(* IEC 61131-3 sources: PLC_I/plc/tests, 6 files *)

(* ---- 程序_气缸自测.st ---- *)
(* 离线IEC扫描自测：放入周期任务，等待b完成，w失败=0才通过。
   不连接物理输出。TON时间证据要求在目标PLC/官方模拟运行，源码测试不能替代。 *)
PROGRAM 程序_气缸自测
VAR
    fb : 功能块_气缸;
    fb原点 : 功能块_气缸;
    ui阶段 : UINT;
    w失败 : WORD;
    b完成 : BOOL;
    t等待 : TON;
    st配置 : 结构体_配置;
    fb调度 : 功能块_气缸调度;
    st运行时 : 结构体_运行时;
    lw原绑定 : LWORD;
    i : UINT;
    udi夹紧请求号 : UDINT; (* 业务示例：保存 Cy动点(Cy夹紧) 返回值 *)
END_VAR
CASE ui阶段 OF
0:
    fb(Execute := FALSE, Token := 0, Code := 0, HasWorkSensor := FALSE, HasOriginSensor := FALSE,
        DelayMs := 20, HomeDelayMs := 30, TimeoutMs := 500, ValveType := 3, HardEstop := FALSE, CancelMode := 0);
    IF fb.AtWork OR fb.AtOrigin OR (fb.DoneToken <> 0) THEN w失败 := 1; END_IF;
    ui阶段 := 1;
1:
    fb(Execute := TRUE, Token := 1, Code := 40);
    IF NOT fb.WorkOutput OR fb.OriginOutput THEN w失败 := 2; END_IF;
    IF fb.DoneToken = 1 THEN ui阶段 := 2; END_IF;
2:
    (* Execute连续TRUE，下一扫描新token仍触发反向请求。 *)
    fb(Execute := TRUE, Token := 2, Code := 41);
    IF fb.WorkOutput OR NOT fb.OriginOutput OR fb.AtWork OR (fb.DoneToken <> 0) THEN w失败 := 3; END_IF;
    ui阶段 := 3;
3:
    fb(Execute := FALSE);
    IF fb.DoneToken = 2 THEN
        IF fb.OriginOutput OR NOT fb.AtOrigin THEN w失败 := 4; END_IF;
        ui阶段 := 4;
    END_IF;
4:
    fb(Execute := TRUE, Token := 3, Code := 40);
    ui阶段 := 5;
5:
    fb(Execute := FALSE, CancelMode := 1);
    IF NOT fb.WorkOutput OR fb.Moving OR fb.AtWork OR fb.AtOrigin OR (fb.DoneToken <> 0) THEN w失败 := 5; END_IF;
    ui阶段 := 6;
6:
    fb(CancelMode := 0);
    IF fb.Moving OR fb.AtWork OR (fb.DoneToken <> 0) THEN w失败 := 6; END_IF;
    ui阶段 := 7;
7:
    fb(Execute := TRUE, Token := 4, Code := 42);
    IF fb.WorkOutput OR fb.OriginOutput OR (fb.DoneToken <> 0) THEN w失败 := 7; END_IF;
    fb原点(Execute := TRUE, Token := 1, Code := 41, HasWorkSensor := FALSE, HasOriginSensor := FALSE,
        DelayMs := 20, HomeDelayMs := 30, TimeoutMs := 500, ValveType := 0, HardEstop := FALSE, CancelMode := 0);
    IF NOT fb原点.Moving OR fb原点.WorkOutput OR fb原点.OriginOutput THEN w失败 := 8; END_IF;
    ui阶段 := 8;
8:
    fb原点(Execute := FALSE);
    IF fb原点.DoneToken = 1 THEN ui阶段 := 9; END_IF;
9:
    fb(Execute := TRUE, Token := 5, Code := 41, CancelMode := 0);
    ui阶段 := 10;
10:
    fb(Execute := FALSE, CancelMode := 1);
    IF fb.OriginOutput OR fb.Moving OR (fb.DoneToken <> 0) THEN w失败 := 9; END_IF;
    ui阶段 := 11;
11:
    fb(Execute := TRUE, Token := 6, Code := 40, CancelMode := 0, HasWorkSensor := TRUE,
        HasOriginSensor := TRUE, SensorWork := TRUE, SensorOrigin := FALSE);
    ui阶段 := 12;
12:
    (* 传感器跌落应重置连续确认延时。 *)
    fb(Execute := FALSE, SensorWork := FALSE);
    IF fb.AtWork OR (fb.DoneToken <> 0) THEN w失败 := 10; END_IF;
    ui阶段 := 13;
13:
    fb(SensorWork := TRUE);
    IF fb.DoneToken = 6 THEN ui阶段 := 14; END_IF;
14:
    fb(HardEstop := TRUE);
    IF NOT fb.Fault OR fb.WorkOutput OR fb.OriginOutput OR (fb.DoneToken <> 0) THEN w失败 := 11; END_IF;
    ui阶段 := 15;
15:
    fb(HardEstop := FALSE);
    IF NOT fb.Fault THEN w失败 := 12; END_IF;
    ui阶段 := 16;
16:
    fb(Execute := TRUE, Token := 7, Code := 42);
    IF fb.Fault OR fb.WorkOutput OR fb.OriginOutput OR (fb.DoneToken <> 0) THEN w失败 := 13; END_IF;
    ui阶段 := 17;
17:
    (* 释放动作未见原点：超时应立即关破真空，不能等待下扫描。 *)
    fb(Execute := TRUE, Token := 8, Code := 41, SensorWork := FALSE, SensorOrigin := FALSE,
        DelayMs := 0, HomeDelayMs := 0, TimeoutMs := 40);
    IF NOT fb.OriginOutput THEN w失败 := 14; END_IF;
    ui阶段 := 18;
18:
    fb(Execute := FALSE);
    IF fb.Fault THEN
        IF (fb.Error <> 2140) OR fb.OriginOutput OR fb.WorkOutput OR fb.Moving THEN w失败 := 15; END_IF;
        ui阶段 := 19;
    END_IF;
19:
    fb(Execute := TRUE, Token := 9, Code := 42);
    fb(Execute := TRUE, Token := 10, Code := 41);
    IF NOT fb.OriginOutput THEN w失败 := 16; END_IF;
    ui阶段 := 20;
20:
    (* 释放中的双传感器冲突同样关破真空。 *)
    fb(Execute := FALSE, SensorWork := TRUE, SensorOrigin := TRUE);
    IF NOT fb.Fault OR (fb.Error <> 2110) OR fb.OriginOutput THEN w失败 := 17; END_IF;
    ui阶段 := 21;
21:
    fb(Execute := TRUE, Token := 11, Code := 42, SensorWork := FALSE, SensorOrigin := FALSE);
    fb(Execute := TRUE, Token := 12, Code := 40);
    ui阶段 := 22;
22:
    (* 吸附超时保持原吸附输出，但绝不打开破真空。 *)
    fb(Execute := FALSE);
    IF fb.Fault THEN
        IF (fb.Error <> 2140) OR NOT fb.WorkOutput OR fb.OriginOutput THEN w失败 := 18; END_IF;
        ui阶段 := 23;
    END_IF;
23:
    (* 独立配置调用：DO0/DI0允许跨空间重号，同空间跨缸别名拒绝。 *)
    lw原绑定 := lw已绑定气缸;
    lw已绑定气缸 := 3;
    FOR i := 0 TO 1 DO
        st配置.aw气缸配置[i, 0] := 0;
        st配置.aw气缸配置[i, 1] := UINT_TO_WORD(i);
        st配置.aw气缸配置[i, 2] := WORD#16#FFFF;
        st配置.aw气缸配置[i, 3] := UINT_TO_WORD(1 - i);
        st配置.aw气缸配置[i, 4] := WORD#16#FFFF;
        st配置.aw气缸配置[i, 5] := 10;
        st配置.aw气缸配置[i, 6] := 100;
        st配置.aw气缸配置[i, 7] := 10;
    END_FOR;
    IF NOT 气缸_配置有效(缸号 := 0, Store := st配置) THEN w失败 := 19; END_IF;
    st配置.aw气缸配置[1, 1] := 0;
    IF 气缸_配置有效(缸号 := 0, Store := st配置) THEN w失败 := 20; END_IF;
    st配置.aw气缸配置[1, 1] := 1;
    st配置.aw气缸配置[1, 3] := 1;
    IF 气缸_配置有效(缸号 := 0, Store := st配置) THEN w失败 := 21; END_IF;
    lw已绑定气缸 := lw原绑定;
    ui阶段 := 24;
24:
    (* 隔离工程中检查真实调度器：手动待复位仍可受理且不被同扫描取消。
       自测不调用物理输出映射，正式工程不得挂此程序。 *)
    lw原绑定 := lw已绑定气缸;
    lw已绑定气缸 := 1;
    FOR i := 0 TO 7 DO
        全局变量_保持区.Store.aw气缸配置[0, i] := st配置.aw气缸配置[0, i];
    END_FOR;
    ab气缸映射有效[0] := TRUE;
    ab气缸模块就绪[0] := TRUE;
    ab气缸动点传感器[0] := FALSE;
    ab气缸原点传感器[0] := FALSE;
    st运行时.b手动 := TRUE;
    st运行时.bHMI在线 := TRUE;
    st运行时.b待复位 := TRUE;
    全局变量_气缸请求.ast请求[0].b自动 := FALSE;
    全局变量_气缸请求.ast请求[0].b待下发 := TRUE;
    全局变量_气缸请求.ast请求[0].b忙 := TRUE;
    全局变量_气缸请求.ast请求[0].udi请求号 := 1;
    全局变量_气缸请求.ast请求[0].w命令 := 40;
    fb调度(StopAll := FALSE, Runtime := st运行时);
    IF NOT ab气缸动点输出[0] OR NOT st运行时.ast气缸[0].b运动中
        OR NOT 全局变量_气缸请求.ast请求[0].b忙 THEN w失败 := 22; END_IF;
    (* 同样待复位条件下自动请求被撤销，不能沿用手动的输出完成资格。 *)
    st运行时.b手动 := FALSE;
    st运行时.b运行 := TRUE;
    全局变量_气缸请求.ast请求[0].b自动 := TRUE;
    全局变量_气缸请求.ast请求[0].b待下发 := TRUE;
    全局变量_气缸请求.ast请求[0].udi请求号 := 2;
    fb调度(StopAll := FALSE, Runtime := st运行时);
    IF st运行时.ast气缸[0].b运动中 OR 全局变量_气缸请求.ast请求[0].b忙 THEN w失败 := 23; END_IF;
    (* 真实语义API：取消覆盖忙槽并登记新令牌；被拒绝动作保留该令牌。 *)
    全局变量_气缸请求.ast请求[0].b忙 := TRUE;
    全局变量_气缸请求.ast请求[0].b待下发 := TRUE;
    IF NOT Cy取消(0) THEN w失败 := 24; END_IF;
    udi夹紧请求号 := Cy设备状态[0].udi请求号;
    IF (udi夹紧请求号 = 0)
        OR (udi夹紧请求号 <> 全局变量_气缸请求.ast请求[0].udi请求号)
        OR (全局变量_气缸请求.ast请求[0].w命令 <> 42) THEN w失败 := 25; END_IF;
    IF Cy动点(0) OR Cy原点(0) THEN w失败 := 26; END_IF;
    IF Cy设备状态[0].udi请求号 <> udi夹紧请求号 THEN w失败 := 27; END_IF;
    IF Cy取消(54) OR Cy动点(54) OR Cy原点(54) THEN w失败 := 28; END_IF;
    lw已绑定气缸 := lw原绑定;
    b完成 := TRUE;
END_CASE;
END_PROGRAM

(* ---- 程序_移植自测.st ---- *)
(* 移植块的行为自测：功能块_输入滤波 / 功能块_运行控制 / 功能块_暂停恢复。
   纯逻辑，不调用 MC，不写物理输出，在隔离仿真器中运行。

   暂停恢复用独立实例、显式输入直接驱动，不经运行状态机：
   每个断言的因果都落在同一个块内，不依赖两个块之间的扫描时序。
   停稳时间用 di停稳ms 参数化，自测取 10 ms，现场仍是 300 ms。 *)
PROGRAM 程序_移植自测
VAR
    fb滤波 : 功能块_输入滤波;
    fb运行 : 功能块_运行控制;
    fb暂停 : 功能块_暂停恢复;
    st运行时 : 结构体_运行时;
    ui阶段 : UINT;
    i循环 : UINT;
    b正常 : BOOL;
    b检查 : BOOL;
    b等待中 : BOOL;
    b首次进入 : BOOL;
    b恢复请求脉冲已发 : BOOL;
    tmr等待 : TON;
    udi通过 : UDINT;
    udi失败 : UDINT;
    ui首失败 : UINT;
    b完成 : BOOL;
    b滤波输入 : BOOL;
    (* 暂停恢复的显式驱动输入。 *)
    b暂停请求 : BOOL;
    b恢复请求 : BOOL;
    b急停测试 : BOOL;
    w诊断1 : WORD;
    w诊断2 : WORD;
END_VAR

IF b完成 THEN RETURN; END_IF;
b检查 := FALSE;
b正常 := TRUE;

(* 运行控制每扫描连续调用；暂停恢复由 b暂停请求 / b恢复请求 直接驱动。 *)
fb运行(b初始化完成 := TRUE,
    b系统复位完成 := TRUE,
    b系统复位中 := FALSE,
    b系统复位失败 := FALSE,
    b启动按钮 := FALSE,
    b暂停按钮 := FALSE,
    b启动事件 := st运行时.b启动脉冲,
    b暂停事件 := st运行时.b暂停脉冲,
    b恢复事件 := st运行时.b恢复脉冲,
    b致命报警 := FALSE,
    b急停 := FALSE,
    b暂停报警 := FALSE,
    b预警 := FALSE,
    b暂停恢复中 := FALSE,
    b暂停恢复完成 := FALSE,
    b暂停恢复失败 := FALSE,
    b流程完成 := FALSE);
st运行时.b启动脉冲 := FALSE;
st运行时.b暂停脉冲 := FALSE;
st运行时.b恢复脉冲 := FALSE;

fb暂停(b暂停 := b暂停请求, b请求 := b恢复请求,
    b急停 := b急停测试,
    di容差 := 100, di停稳ms := 10, Runtime := st运行时);

(* 等待解除：条件满足或超时都只做一次“解除 b等待中”，推进交给扫描末尾统一处理。
   这样每个扫描最多推进一次，阶段体不会重复执行，也不会漏推进。 *)
tmr等待(IN := b等待中, PT := T#500ms);
IF b等待中 THEN
    IF (ui阶段 = 10) AND fb暂停.b已抓拍 THEN b等待中 := FALSE;
    ELSIF (ui阶段 = 16) AND (st运行时.aw轴命令[0] = 27) THEN b等待中 := FALSE;
    ELSIF (ui阶段 = 18) AND (fb暂停.b恢复完成 OR fb暂停.b恢复失败) THEN b等待中 := FALSE;
    ELSIF tmr等待.Q THEN b等待中 := FALSE;
    END_IF;
END_IF;
(* b等待中 只由阶段体在“首次进入”时置位，由上面的条件或 500 ms 超时解除；
   扫描末尾按它的值决定是否推进，因此每个扫描最多推进一次。 *)

w诊断1 := fb暂停.ui内部阶段 * 256;
IF fb暂停.b已抓拍 THEN w诊断1 := w诊断1 OR 2; END_IF;
IF fb暂停.b曾偏离 THEN w诊断1 := w诊断1 OR 4; END_IF;
IF fb暂停.b恢复中 THEN w诊断1 := w诊断1 OR 8; END_IF;
IF fb暂停.b恢复完成 THEN w诊断1 := w诊断1 OR 16; END_IF;
IF fb暂停.b恢复失败 THEN w诊断1 := w诊断1 OR 32; END_IF;
w诊断2 := 0;
IF st运行时.aw轴命令[0] = 27 THEN w诊断2 := w诊断2 OR 1; END_IF;
IF st运行时.aw轴命令[0] = 26 THEN w诊断2 := w诊断2 OR 2; END_IF;

CASE ui阶段 OF
    (* ===== 输入滤波 ===== *)
    0:
        b滤波输入 := TRUE;
        fb滤波(b信号 := b滤波输入, i模式 := 0,
            di滤波时间真 := 20, di滤波时间假 := 20);
        b检查 := TRUE; b正常 := fb滤波.b滤波信号;
    1:
        (* 模式 1：输入变 FALSE，20 ms 未到，输出保持上一扫描的 TRUE。 *)
        b滤波输入 := FALSE;
        fb滤波(b信号 := b滤波输入, i模式 := 1,
            di滤波时间真 := 20, di滤波时间假 := 20);
        b检查 := TRUE; b正常 := fb滤波.b滤波信号;
    2:
        (* 非法模式按直通，不把输入锁死。 *)
        b滤波输入 := TRUE;
        fb滤波(b信号 := b滤波输入, i模式 := 99,
            di滤波时间真 := 20, di滤波时间假 := 20);
        b检查 := TRUE; b正常 := fb滤波.b滤波信号;

    (* ===== 运行控制 ===== *)
    3:
        b检查 := TRUE;
        b正常 := fb运行.b手动模式 AND NOT fb运行.b运行指令 AND NOT fb运行.b暂停中;
    4:
        st运行时.b启动脉冲 := TRUE;
    5:
        b检查 := TRUE;
        b正常 := fb运行.b运行指令 AND NOT fb运行.b暂停中 AND fb运行.b自动模式;
    6:
        st运行时.b暂停脉冲 := TRUE;
    7:
        b检查 := TRUE; b正常 := (NOT fb运行.b运行指令) AND fb运行.b暂停中;
    8:
        (* 暂停优先于启动：暂停中收到启动不得运行。 *)
        st运行时.b启动脉冲 := TRUE;
    9:
        b检查 := TRUE; b正常 := (NOT fb运行.b运行指令) AND fb运行.b暂停中;

    (* ===== 暂停恢复：直接驱动 ===== *)
    10:
        (* 三轴静止于 1000，无急停，进入暂停。
           进入后立刻布置等待；阶段体不再重复执行，避免每扫描重置等待。 *)
        IF b首次进入 THEN
        b首次进入 := FALSE;
        b等待中 := TRUE;
        st运行时.w轴消费掩码 := 7;
        st运行时.bHMI在线 := TRUE;
        st运行时.b待复位 := FALSE;
        st运行时.b暂停 := TRUE;
        FOR i循环 := 0 TO 2 DO
            全局变量_保持区.Store.aw轴配置[i循环, 0] := 0;
            全局变量_保持区.Store.aw轴配置[i循环, 1] := 10000;
            全局变量_保持区.Store.aw轴配置[i循环, 2] := WORD#16#FFFF;
            全局变量_保持区.Store.aw轴配置[i循环, 3] := WORD#16#D8F0;
            全局变量_保持区.Store.aw轴配置[i循环, 14] := 1;
            全局变量_保持区.Store.aw轴配置[i循环, 4] := 0;
            全局变量_保持区.Store.aw轴配置[i循环, 5] := 1000;
            全局变量_保持区.Store.aw轴配置[i循环, 6] := 0;
            全局变量_保持区.Store.aw轴配置[i循环, 7] := 1000;
            全局变量_保持区.Store.aw轴配置[i循环, 8] := 0;
            全局变量_保持区.Store.aw轴配置[i循环, 9] := 1000;
            全局变量_保持区.Store.aw轴配置[i循环, 10] := 0;
            全局变量_保持区.Store.aw轴配置[i循环, 11] := 1000;
            全局变量_保持区.Store.aw轴配置[i循环, 12] := 0;
            全局变量_保持区.Store.aw轴配置[i循环, 13] := 1000;
            st运行时.ast轴[i循环].b已使能 := TRUE;
            st运行时.ast轴[i循环].b可下发 := TRUE;
        END_FOR;
        b急停测试 := FALSE;
        b恢复请求 := FALSE;
        FOR i循环 := 0 TO 2 DO
            st运行时.ast轴[i循环].b在线 := TRUE;
            st运行时.ast轴[i循环].b静止 := TRUE;
            st运行时.ast轴[i循环].b运动中 := FALSE;
            st运行时.ast轴[i循环].b故障 := FALSE;
            st运行时.ast轴[i循环].di位置 := 1000;
            st运行时.ast轴[i循环].w序列 := 0;
            st运行时.ast轴[i循环].w运动结果 := 0;
        END_FOR;
        b暂停请求 := TRUE;
        END_IF;
    11:
        (* 停稳 10 ms 后必须抓到快照。 *)
        b检查 := TRUE; b正常 := fb暂停.b已抓拍;
    12:
        (* 未偏离时请求恢复。恢复请求是上升沿事件，置位一个扫描即撤销。 *)
        b恢复请求 := TRUE;
    13:
        b恢复请求 := FALSE;
        b检查 := TRUE;
        b正常 := fb暂停.b恢复完成 AND NOT fb暂停.b恢复失败 AND (st运行时.aw轴命令[0] = 0);
    14:
        (* 拉开轴 0 超出容差 100：应锁存曾偏离。 *)
        b恢复请求 := FALSE;
        st运行时.ast轴[0].di位置 := 2000;
    15:
        b检查 := TRUE; b正常 := fb暂停.b曾偏离;
    16:
        (* 请求恢复：应给轴 0 下发绝对定位 27 回快照位置 1000。 *)
        IF b首次进入 THEN
        b首次进入 := FALSE;
        b等待中 := TRUE;
        st运行时.ast轴[0].w序列 := 0;
        st运行时.ast轴[0].w运动结果 := 0;
        b恢复请求 := TRUE;
        END_IF;
        (* 恢复请求保持到完成，撤销请求将主动停止正在回位的轴。 *)
    17:
        b检查 := TRUE;
        b正常 := (st运行时.aw轴命令[0] = 27) AND (st运行时.adi轴目标[0] = 1000);
    18:
        (* 轴报告结果 2 且静止：恢复完成。 *)
        st运行时.ast轴[0].w序列 := st运行时.aw轴序列[0];
        st运行时.ast轴[0].w运动结果 := 2;
        st运行时.ast轴[0].di位置 := 1000;
        IF b首次进入 THEN
        b首次进入 := FALSE;
        b等待中 := TRUE;
        st运行时.ast轴[0].b静止 := TRUE;
        st运行时.ast轴[0].b运动中 := FALSE;
        END_IF;
    19:
        b检查 := TRUE; b正常 := fb暂停.b恢复完成 AND NOT fb暂停.b恢复失败;
    20:
        (* 急停：必须封锁并撤销本块下发的命令。 *)
        b恢复请求 := FALSE;
        st运行时.ast轴[0].di位置 := 3000;
        st运行时.aw轴命令[0] := 0; (* 服务端每扫描清命令槽 *)
        b急停测试 := TRUE;
    21: ;
    22:
        b检查 := TRUE; b正常 := st运行时.aw轴命令[0] = 0;
    23:
        b急停测试 := FALSE;
        st运行时.aw轴命令[0] := 0;
        st运行时.b待复位 := TRUE;
        b恢复请求 := TRUE;
    24:
        b检查 := TRUE; b正常 := fb暂停.b恢复失败 AND (st运行时.aw轴命令[0] = 0);
        b恢复请求 := FALSE;
        st运行时.b待复位 := FALSE;
        (* 快照1000在新软限位之外，即使其他条件满足仍不得回位。 *)
        全局变量_保持区.Store.aw轴配置[0, 3] := 1500;
        全局变量_保持区.Store.aw轴配置[0, 2] := 0;
    25:
        b恢复请求 := TRUE;
    26:
        b检查 := TRUE; b正常 := fb暂停.b恢复失败 AND (st运行时.aw轴命令[0] = 0);
        b恢复请求 := FALSE;
        全局变量_保持区.Store.aw轴配置[0, 2] := WORD#16#FFFF;
        全局变量_保持区.Store.aw轴配置[0, 3] := WORD#16#D8F0;
    27:
        b恢复请求 := TRUE;
    28:
        b检查 := TRUE; b正常 := st运行时.aw轴命令[0] = 27;
        st运行时.aw轴命令[0] := 0; (* emulate server clearing pulse slot *)
        st运行时.ast轴[0].b运动中 := TRUE;
        st运行时.ast轴[0].b静止 := FALSE;
        st运行时.ast轴[0].b可下发 := FALSE;
    29:
        (* 本动作自身Busy不可被持续复核误判成失许可。 *)
        b检查 := TRUE; b正常 := fb暂停.b恢复中 AND NOT fb暂停.b恢复失败;
        st运行时.bHMI在线 := FALSE;
    30:
        b检查 := TRUE; b正常 := fb暂停.b恢复失败 AND (st运行时.aw轴命令[0] = 26);
        b完成 := TRUE;
END_CASE;

IF b检查 THEN
    IF b正常 THEN udi通过 := udi通过 + 1;
    ELSE
        udi失败 := udi失败 + 1;
        IF ui首失败 = 0 THEN ui首失败 := ui阶段; END_IF;
    END_IF;
END_IF;
(* b等待中 可能在阶段体内刚被置位，这里同时看两个标志，避免立即推进。 *)
(* 每个扫描最多推进一次。阶段体若在本扫描刚置 b等待中，就保持不动。 *)
IF NOT b等待中 THEN ui阶段 := ui阶段 + 1; b首次进入 := TRUE; END_IF;
END_PROGRAM

(* ---- 程序_自测.st ---- *)
(* Isolated simulator test task only. Never schedule with real machine control.
   Cold/reset-origin starts a fresh run; Done latches until the next reset.
   Watch 程序_自测.Passed/Failed/Done/FirstFailure.
   Protocol 1.2: Modbus is the official slave device, so the former Access
   adapter cases are gone; requests are fed to 功能块_配置 directly.
   Expected terminal result: Done=TRUE, Passed=61, Failed=0, FirstFailure=0.
   FirstFailure is the 1-based case ID (Step + 1); one case per active scan,
   separated by an idle scan to release Execute and Request.
   No network, device references, retained GVL, external assertion or library.
*)
PROGRAM 程序_自测
VAR
    udi通过 : UDINT;
    udi失败 : UDINT;
    b完成 : BOOL;
    ui首失败 : UINT;
    ui首失败步骤 : UINT;
    w首失败结果 : WORD;
    w首失败对象 : WORD;
    ui步骤 : UINT;
    b空闲扫描 : BOOL;
    fb配置 : 功能块_配置;
    st配置 : 结构体_配置;
    st原配置 : 结构体_配置;
    st请求 : 类型_命令区;
    w原纪元 : WORD;
    w原结果 : WORD;
    w期望纪元 : WORD;
    w期望结果 : WORD;
    b执行配置 : BOOL;
    b检查回滚 : BOOL;
    b检查空闲 : BOOL;
    b正常 : BOOL;
    i点位索引 : INT;
    i循环 : INT;
    i子循环 : INT;
END_VAR

IF b完成 THEN RETURN; END_IF;
IF b空闲扫描 THEN
    fb配置(Execute := FALSE, Request := st请求, Store := st配置);
    b空闲扫描 := FALSE;
    RETURN;
END_IF;

FOR i循环 := 0 TO 31 DO st请求[i循环] := 0; END_FOR;
st请求[0] := WORD#16#584A;
st请求[1] := XJV1_SIGNATURE_LO;
st请求[4] := 1;
st请求[5] := WORD#16#0100;
b执行配置 := FALSE;
b检查回滚 := FALSE;
b检查空闲 := FALSE;
w期望结果 := 0;
b正常 := TRUE;

CASE ui步骤 OF
    0:
        st配置.dw签名 := 0;
        st配置.b已确认 := TRUE;
    1:
        (* Wrong signature is rejected before any record changes. *)
        st请求[1] := WORD#16#5631; st请求[3] := 31; st请求[7] := 19; st请求[11] := 1;
        b执行配置 := TRUE; b检查回滚 := TRUE; w期望结果 := 1;
    2:
        (* Non-zero reserved header word +15. *)
        st请求[3] := 31; st请求[7] := 19; st请求[11] := 1; st请求[15] := 1;
        b执行配置 := TRUE; b检查回滚 := TRUE; w期望结果 := 9;
    3:
        (* Command 51 (retired PLC name commit) is unsupported. *)
        st请求[3] := 51; st请求[5] := WORD#16#0100;
        b执行配置 := TRUE; b检查回滚 := TRUE; w期望结果 := 14;
    4:
        (* Code 50 on the system object is an illegal object. *)
        st请求[3] := 50; st请求[5] := 0; st请求[7] := 1;
        b执行配置 := TRUE; b检查回滚 := TRUE; w期望结果 := 15;
    5:
        (* Point index 120 is out of the pool. *)
        st请求[3] := 50; st请求[5] := WORD#16#0378; st请求[7] := 4;
        b执行配置 := TRUE; b检查回滚 := TRUE; w期望结果 := 15;
    6:
        (* Free slots are exactly XJV1_POINT_FREE after cold init. *)
        b检查空闲 := TRUE; b检查回滚 := TRUE;
        b正常 := (st配置.aw点位[19, 4] = XJV1_POINT_FREE) AND (fb配置.Epoch = 0);
    7:
        (* Free bit combined with an owner is never accepted. *)
        st请求[3] := 50; st请求[5] := WORD#16#0313; st请求[7] := 4; st请求[9] := fb配置.Epoch;
        FOR i循环 := 0 TO 4 DO st请求[16 + i循环] := st配置.aw点位[19, i循环]; END_FOR;
        st请求[20] := XJV1_POINT_FREE OR WORD#16#0004;
        b执行配置 := TRUE; b检查回滚 := TRUE; w期望结果 := 9;
    8:
        (* Release of P0 standby slot 0 (owned by axis 0) is rejected. *)
        st请求[3] := 50; st请求[5] := WORD#16#0300; st请求[7] := 4; st请求[9] := fb配置.Epoch;
        FOR i循环 := 0 TO 4 DO st请求[16 + i循环] := st配置.aw点位[0, i循环]; END_FOR;
        st请求[20] := XJV1_POINT_FREE;
        b执行配置 := TRUE; b检查回滚 := TRUE; w期望结果 := 9;
    9:
        (* Stale config epoch. *)
        st请求[3] := 50; st请求[5] := WORD#16#0313; st请求[7] := 4; st请求[9] := fb配置.Epoch + 1;
        FOR i循环 := 0 TO 4 DO st请求[16 + i循环] := st配置.aw点位[19, i循环]; END_FOR;
        st请求[20] := WORD#16#0000;
        b执行配置 := TRUE; b检查回滚 := TRUE; w期望结果 := 16;
    10:
        (* Teach claims free slot 19 for axis 0: position -1000, speed 65536. *)
        st请求[3] := 31; st请求[7] := 19;
        st请求[8] := WORD#16#FFFF; st请求[9] := WORD#16#FC18;
        st请求[10] := 1; st请求[11] := 0;
        b执行配置 := TRUE;
    11:
        st请求[3] := 31; st请求[7] := 19; st请求[11] := 1; st请求[15] := 1;
        b执行配置 := TRUE; b检查回滚 := TRUE; w期望结果 := 9;
    12..31:
        i点位索引 := UINT_TO_INT(ui步骤) - 12;
        (* Deliberate fixture: alternating disabled/enabled already-taught points. *)
        IF (i点位索引 MOD 2) = 0 THEN st配置.aw点位[i点位索引, 4] := 0;
        ELSE st配置.aw点位[i点位索引, 4] := 3; END_IF;
        st配置.b已确认 := TRUE;
        st请求[3] := 31;
        st请求[7] := INT_TO_WORD(i点位索引);
        st请求[8] := WORD#16#FFFF;
        st请求[9] := DINT_TO_WORD(DINT#64536 - INT_TO_DINT(i点位索引));
        st请求[10] := 1; st请求[11] := INT_TO_WORD(i点位索引);
        b执行配置 := TRUE;
    32..37:
        st请求[3] := 50;
        st请求[7] := 4;
        st请求[9] := fb配置.Epoch;
        FOR i循环 := 0 TO 15 DO st请求[16 + i循环] := st配置.aw轴配置[0, i循环]; END_FOR;
        b执行配置 := TRUE;
        CASE ui步骤 OF
            32:
                st配置.b已确认 := TRUE;
                st请求[16] := 0; st请求[17] := 0;
                st请求[20] := 1; st请求[21] := 2;
            33:
                st请求[20] := 0; st请求[21] := 0;
                b检查回滚 := TRUE; w期望结果 := 22;
            34:
                st请求[7] := 1;
                st请求[16] := st配置.aw轴配置[0, 2]; st请求[17] := st配置.aw轴配置[0, 3];
                b检查回滚 := TRUE; w期望结果 := 21;
            35:
                st请求[9] := 0;
                b检查回滚 := TRUE; w期望结果 := 16;
            36:
                st请求[8] := 1;
                b检查回滚 := TRUE; w期望结果 := 9;
            37:
                st请求[31] := 1;
                b检查回滚 := TRUE; w期望结果 := 9;
        END_CASE;
    38:
        st请求[3] := 50; st请求[5] := WORD#16#0314;
        st请求[7] := 4; st请求[9] := fb配置.Epoch;
        FOR i循环 := 0 TO 4 DO st请求[16 + i循环] := st配置.aw点位[20, i循环]; END_FOR;
        st请求[20] := 3;
        b执行配置 := TRUE; b检查回滚 := TRUE; w期望结果 := 9;
    39:
        st配置.aw点位[19, 4] := 2;
        st配置.b已确认 := TRUE;
        st请求[3] := 50; st请求[5] := WORD#16#0313;
        st请求[7] := 4; st请求[9] := fb配置.Epoch;
        FOR i循环 := 0 TO 4 DO st请求[16 + i循环] := st配置.aw点位[19, i循环]; END_FOR;
        st请求[20] := 3;
        b执行配置 := TRUE;
    40:
        st请求[3] := 31; st请求[7] := 19;
        st请求[8] := WORD#16#8000; st请求[9] := 0;
        st请求[10] := WORD#16#7FFF; st请求[11] := WORD#16#FFFF;
        b执行配置 := TRUE;
    41..50:
        (* Retired name commit 51 must stay unsupported for every object kind. *)
        st请求[3] := 51;
        CASE ui步骤 OF
            41, 42, 43: st请求[5] := WORD#16#0100;
            44, 45, 46: st请求[5] := WORD#16#0200;
        ELSE st请求[5] := WORD#16#0300;
        END_CASE;
        st请求[7] := fb配置.Epoch; st请求[16] := 65;
        b执行配置 := TRUE; b检查回滚 := TRUE; w期望结果 := 14;
    51..53:
        st请求[3] := 31; st请求[7] := 19; st请求[11] := 1;
        b执行配置 := TRUE; b检查回滚 := TRUE; w期望结果 := 9;
        CASE ui步骤 OF
            51: st请求[6] := 1;
            52: st请求[7] := 120;
            53: st请求[10] := WORD#16#8000; st请求[11] := 0;
        END_CASE;
    54:
        b检查空闲 := TRUE; b检查回滚 := TRUE;
    55:
        (* Cylinder 1 is unbound in production binding: parameter commit rejects 4. *)
        st请求[3] := 50; st请求[5] := WORD#16#0201; st请求[7] := 1; st请求[9] := fb配置.Epoch;
        FOR i循环 := 0 TO 7 DO st请求[16 + i循环] := st配置.aw气缸配置[1, i循环]; END_FOR;
        b执行配置 := TRUE; b检查回滚 := TRUE; w期望结果 := 4;
    56:
        (* Axis 15 owner bits (16#003C) and the free code are distinct. Slot 15's
           cold-init owner is verified in step 0; slots 0..19 are re-owned by the
           step 12..31 fixture, so check an untouched free slot here. *)
        b检查空闲 := TRUE; b检查回滚 := TRUE;
        b正常 := (st配置.aw点位[20, 4] = XJV1_POINT_FREE) AND (XJV1_POINT_FREE <> SHL(WORD#15, 2));
    57:
        (* Point index 160 is out of range. *)
        st请求[3] := 50; st请求[5] := WORD#16#03A0; st请求[7] := 4;
        b执行配置 := TRUE; b检查回滚 := TRUE; w期望结果 := 15;
    58:
        st请求[3] := 50; st请求[5] := WORD#16#0313;
        st请求[7] := 2; st请求[9] := fb配置.Epoch;
        FOR i循环 := 0 TO 4 DO st请求[16 + i循环] := st配置.aw点位[19, i循环]; END_FOR;
        st请求[18] := WORD#16#8000; st请求[19] := 0;
        b执行配置 := TRUE; b检查回滚 := TRUE; w期望结果 := 9;
    59:
        (* Release slot 19: disable + untaught is required; taught slot rejects 9. *)
        st请求[3] := 50; st请求[5] := WORD#16#0313; st请求[7] := 4; st请求[9] := fb配置.Epoch;
        FOR i循环 := 0 TO 4 DO st请求[16 + i循环] := st配置.aw点位[19, i循环]; END_FOR;
        st请求[20] := XJV1_POINT_FREE;
        b执行配置 := TRUE; b检查回滚 := TRUE; w期望结果 := 9;
    60:
        st请求[3] := 31; st请求[7] := 19; st请求[11] := 999;
        b检查空闲 := TRUE; b检查回滚 := TRUE;
ELSE
    b正常 := FALSE;
END_CASE;

st原配置 := st配置;
w原纪元 := fb配置.Epoch;
w原结果 := fb配置.Result;
fb配置(Execute := b执行配置, Request := st请求, Store := st配置);
IF b执行配置 THEN
    IF fb配置.Result <> w期望结果 THEN b正常 := FALSE; END_IF;
    w期望纪元 := w原纪元;
    IF w期望结果 = 0 THEN
        IF w原纪元 = WORD#16#FFFF THEN w期望纪元 := 0;
        ELSE w期望纪元 := w原纪元 + 1; END_IF;
    END_IF;
    IF fb配置.Epoch <> w期望纪元 THEN b正常 := FALSE; END_IF;
END_IF;
IF b检查空闲 AND (fb配置.Result <> w原结果) THEN b正常 := FALSE; END_IF;

IF b检查回滚 THEN
    IF (fb配置.Epoch <> w原纪元) OR (st配置.dw签名 <> st原配置.dw签名)
    OR (st配置.b已确认 <> st原配置.b已确认) THEN b正常 := FALSE; END_IF;
    FOR i循环 := 0 TO 15 DO
        FOR i子循环 := 0 TO 15 DO
            IF st配置.aw轴配置[i循环, i子循环] <> st原配置.aw轴配置[i循环, i子循环] THEN b正常 := FALSE; END_IF;
        END_FOR;
    END_FOR;
    FOR i循环 := 0 TO 53 DO
        FOR i子循环 := 0 TO 7 DO
            IF st配置.aw气缸配置[i循环, i子循环] <> st原配置.aw气缸配置[i循环, i子循环] THEN b正常 := FALSE; END_IF;
        END_FOR;
    END_FOR;
    FOR i循环 := 0 TO 119 DO
        FOR i子循环 := 0 TO 4 DO
            IF st配置.aw点位[i循环, i子循环] <> st原配置.aw点位[i循环, i子循环] THEN b正常 := FALSE; END_IF;
        END_FOR;
    END_FOR;
END_IF;

CASE ui步骤 OF
    0:
        b正常 := (st配置.dw签名 = XJV1_SIGNATURE) AND NOT st配置.b已确认 AND (fb配置.Epoch = 0);
        FOR i循环 := 0 TO 119 DO
            IF i循环 < 16 THEN
                IF st配置.aw点位[i循环, 4] <> SHL(INT_TO_WORD(i循环), 2) THEN b正常 := FALSE; END_IF;
            ELSIF st配置.aw点位[i循环, 4] <> XJV1_POINT_FREE THEN b正常 := FALSE; END_IF;
            IF st配置.aw点位[i循环, 3] <> 1 THEN b正常 := FALSE; END_IF;
        END_FOR;
        FOR i循环 := 0 TO 53 DO
            FOR i子循环 := 1 TO 4 DO
                IF st配置.aw气缸配置[i循环, i子循环] <> WORD#16#FFFF THEN b正常 := FALSE; END_IF;
            END_FOR;
            IF (st配置.aw气缸配置[i循环, 5] <> 200) OR (st配置.aw气缸配置[i循环, 6] <> 3000) THEN b正常 := FALSE; END_IF;
        END_FOR;
    10:
        IF (st配置.aw点位[19, 0] <> WORD#16#FFFF) OR (st配置.aw点位[19, 1] <> WORD#16#FC18)
        OR (st配置.aw点位[19, 2] <> 1) OR (st配置.aw点位[19, 3] <> 0)
        OR (st配置.aw点位[19, 4] <> 2) OR st配置.b已确认 THEN b正常 := FALSE; END_IF;
    12..31:
        IF (st配置.aw点位[i点位索引, 0] <> WORD#16#FFFF)
        OR (st配置.aw点位[i点位索引, 1] <> DINT_TO_WORD(DINT#64536 - INT_TO_DINT(i点位索引)))
        OR (st配置.aw点位[i点位索引, 2] <> 1) OR (st配置.aw点位[i点位索引, 3] <> INT_TO_WORD(i点位索引))
        OR (st配置.aw点位[i点位索引, 4] <> (st原配置.aw点位[i点位索引, 4] OR WORD#16#0002))
        OR st配置.b已确认 THEN b正常 := FALSE; END_IF;
    32:
        FOR i子循环 := 0 TO 15 DO
            IF i子循环 = 4 THEN
                IF st配置.aw轴配置[0, i子循环] <> 1 THEN b正常 := FALSE; END_IF;
            ELSIF i子循环 = 5 THEN
                IF st配置.aw轴配置[0, i子循环] <> 2 THEN b正常 := FALSE; END_IF;
            ELSIF st配置.aw轴配置[0, i子循环] <> st原配置.aw轴配置[0, i子循环] THEN b正常 := FALSE;
            END_IF;
        END_FOR;
        IF st配置.b已确认 THEN b正常 := FALSE; END_IF;
    39:
        IF (st配置.aw点位[19, 4] <> 3) OR st配置.b已确认 THEN b正常 := FALSE; END_IF;
        FOR i子循环 := 0 TO 3 DO
            IF st配置.aw点位[19, i子循环] <> st原配置.aw点位[19, i子循环] THEN b正常 := FALSE; END_IF;
        END_FOR;
    40:
        IF (st配置.aw点位[19, 0] <> WORD#16#8000) OR (st配置.aw点位[19, 1] <> 0)
        OR (st配置.aw点位[19, 2] <> WORD#16#7FFF) OR (st配置.aw点位[19, 3] <> WORD#16#FFFF)
        OR (st配置.aw点位[19, 4] <> 3) THEN b正常 := FALSE; END_IF;
END_CASE;

IF b正常 THEN
    udi通过 := udi通过 + 1;
ELSE
    udi失败 := udi失败 + 1;
    IF ui首失败 = 0 THEN ui首失败 := ui步骤 + 1; END_IF;
    IF ui首失败 = ui步骤 + 1 THEN
        ui首失败步骤 := ui步骤;
        w首失败结果 := fb配置.Result;
        w首失败对象 := st请求[5];
    END_IF;
END_IF;
IF ui步骤 >= 60 THEN
    b完成 := TRUE;
ELSE
    ui步骤 := ui步骤 + 1;
    b空闲扫描 := TRUE;
END_IF;
END_PROGRAM

(* ---- 程序_轴报警自测.st ---- *)
(* Offline adapter behavior with mock MC blocks. Never run on physical axes. *)
PROGRAM PRG_AxisAlarmTest
VAR
    Step : UINT;
    Passed : UINT;
    Failed : UINT;
    Done : BOOL;
    DummyAxis : AXIS_REF_SM3;
    Motion : FB_AxisUnderTest;
    Fault : FB_AxisUnderTest;
    InvalidRead : FB_AxisUnderTest;
    FailedRead : FB_AxisUnderTest;
    Bus : FB_AxisUnderTest;
    Emergency : FB_AxisUnderTest;
    Pulse : FB_AxisUnderTest;
    States : ARRAY[0..5] OF 结构体_轴状态;
    PulseState : 结构体_轴状态;
    LimitStop : FB_AxisUnderTest;
    SoftwareStop : FB_AxisUnderTest;
    LimitState : 结构体_轴状态;
    SoftwareState : 结构体_轴状态;
END_VAR

CASE Step OF
0:
    Motion(Axis := DummyAxis, State := States[0], Code := 0);
    Fault(Axis := DummyAxis, State := States[1], Code := 0);
    InvalidRead(Axis := DummyAxis, State := States[2], Code := 0);
    FailedRead(Axis := DummyAxis, State := States[3], Code := 0);
    Bus(Axis := DummyAxis, State := States[4], Code := 0, BusOperational := FALSE);
    Emergency(Axis := DummyAxis, State := States[5], Code := 0);
    Pulse.fb读位置.Valid := FALSE;
    Pulse.fb读速度.Valid := FALSE;
    Pulse(Axis := DummyAxis, State := PulseState, Code := 0, OpenLoop := TRUE);
    IF PulseState.b在线 AND NOT PulseState.b已使能 THEN Passed := Passed + 1;
    ELSE Failed := Failed + 1; END_IF;
    IF States[0].b在线 AND NOT States[4].b在线 THEN Passed := Passed + 1;
    ELSE Failed := Failed + 1; END_IF;
    Step := 1;
1:
    Motion(Axis := DummyAxis, State := States[0], Code := 20, Sequence := 1);
    Step := 2;
2:
    Motion(Axis := DummyAxis, State := States[0], Code := 24, Sequence := 2,
        Speed := 5000, Acceleration := 2000, Deceleration := 3000, StopDeceleration := 0);
    IF Motion.lr锁定停止减速度 = 3.0 AND States[0].b正向点动 THEN Passed := Passed + 1;
    ELSE Failed := Failed + 1; END_IF;
    Fault.fb读状态.Errorstop := TRUE;
    Fault.fb读轴错.AxisErrorID := DWORD#16#1234;
    Fault(Axis := DummyAxis, State := States[1], Code := 0);
    IF (States[1].w错误码 = 1104) AND (States[1].dw驱动错误 = DWORD#16#1234) THEN Passed := Passed + 1;
    ELSE Failed := Failed + 1; END_IF;
    IF NOT Fault.fb上电.Enable THEN Passed := Passed + 1;
    ELSE Failed := Failed + 1; END_IF;
    InvalidRead.fb读状态.Errorstop := TRUE;
    InvalidRead.fb读轴错.Valid := FALSE;
    InvalidRead.fb读轴错.AxisErrorID := DWORD#16#1234;
    InvalidRead(Axis := DummyAxis, State := States[2], Code := 0);
    IF (States[2].w错误码 = 1104) AND (States[2].dw驱动错误 = 0) THEN Passed := Passed + 1;
    ELSE Failed := Failed + 1; END_IF;
    FailedRead.fb读状态.Errorstop := TRUE;
    FailedRead.fb读轴错.Valid := FALSE;
    FailedRead.fb读轴错.Error := TRUE;
    FailedRead.fb读轴错.ErrorID := DWORD#16#55;
    FailedRead.fb读轴错.AxisErrorID := DWORD#16#1234;
    FailedRead(Axis := DummyAxis, State := States[3], Code := 0);
    IF (States[3].w错误码 = 1104) AND (States[3].dw驱动错误 = DWORD#16#55) THEN Passed := Passed + 1;
    ELSE Failed := Failed + 1; END_IF;
    Bus(Axis := DummyAxis, State := States[4], Code := 20, BusOperational := FALSE);
    IF NOT States[4].b在线 AND NOT States[4].b已使能 THEN Passed := Passed + 1;
    ELSE Failed := Failed + 1; END_IF;
    Emergency(Axis := DummyAxis, State := States[5], Code := 20, HardEstop := TRUE);
    IF (States[5].w错误码 = 1103) AND NOT States[5].b已使能 THEN Passed := Passed + 1;
    ELSE Failed := Failed + 1; END_IF;
    Step := 3;
3:
    Fault(Axis := DummyAxis, State := States[1], Code := 23, Sequence := 3);
    IF Fault.fb复位.Execute AND NOT Fault.fb上电.Enable THEN Passed := Passed + 1;
    ELSE Failed := Failed + 1; END_IF;
    LimitStop(Axis := DummyAxis, State := LimitState, Code := 0);
    SoftwareStop(Axis := DummyAxis, State := SoftwareState, Code := 0);
    Step := 4;
4:
    LimitStop(Axis := DummyAxis, State := LimitState, Code := 20, Sequence := 1);
    SoftwareStop(Axis := DummyAxis, State := SoftwareState, Code := 20, Sequence := 1);
    Fault.fb复位.Done := TRUE;
    Fault.fb读状态.Errorstop := FALSE;
    Fault(Axis := DummyAxis, State := States[1], Code := 0);
    IF NOT Fault.b请求上电 AND NOT States[1].b已使能 AND NOT States[1].b故障 THEN Passed := Passed + 1;
    ELSE Failed := Failed + 1; END_IF;
    Step := 5;
5:
    LimitStop(Axis := DummyAxis, State := LimitState, Code := 27, Sequence := 2,
        Target := 10000, Speed := 5000, Acceleration := 2000, Deceleration := 3000);
    SoftwareStop(Axis := DummyAxis, State := SoftwareState, Code := 27, Sequence := 2,
        Target := 10000, Speed := 5000, Acceleration := 2000, Deceleration := 3000);
    Step := 6;
6:
    LimitStop.fb读状态.StandStill := FALSE;
    LimitStop.fb读状态.DiscreteMotion := TRUE;
    LimitStop.fb读速度.Velocity := 1.0;
    LimitStop(Axis := DummyAxis, State := LimitState, Code := 0, PositiveLimit := TRUE);
    IF LimitStop.fb停止.Execute AND NOT LimitStop.b执行运动 AND (LimitStop.w激活命令 = 0) THEN Passed := Passed + 1;
    ELSE Failed := Failed + 1; END_IF;
    SoftwareStop.fb读状态.StandStill := FALSE;
    SoftwareStop.fb读状态.DiscreteMotion := TRUE;
    SoftwareStop.fb读速度.Velocity := 1.0;
    SoftwareStop.fb读位置.Position := LREAL#3000000; (* conversion fault while physically moving *)
    SoftwareStop(Axis := DummyAxis, State := SoftwareState, Code := 0);
    (* Position invalid prevents MC_Stop: power must be removed rather than leave motion enabled. *)
    IF SoftwareState.b故障 AND NOT SoftwareStop.b请求上电 THEN Passed := Passed + 1;
    ELSE Failed := Failed + 1; END_IF;
    Step := 7;
7:
    (* 软件报警本身不能阻止有效驱动制动。 *)
    LimitState.b故障 := TRUE;
    LimitStop(Axis := DummyAxis, State := LimitState, Code := 0);
    IF LimitStop.fb停止.Execute AND LimitStop.b请求上电 THEN Passed := Passed + 1;
    ELSE Failed := Failed + 1; END_IF;
    Done := TRUE;
    Step := 8;
END_CASE;
END_PROGRAM

(* ---- 程序_轴接口自测.st ---- *)
(* Isolated logic test: real API and server, synthetic axis feedback, no MC/IO. *)
PROGRAM 程序_轴接口自测
VAR
    Server : 功能块_服务端;
    Manager : 功能块_轴请求监视;
    Runtime : 结构体_运行时;
    Command : 类型_命令区;
    Published : 类型_发布区;
    Step : UINT;
    Passed : UDINT;
    Failed : UDINT;
    FirstFailure : UINT;
    Done : BOOL;
    Ok : BOOL;
    Check : BOOL;
    Result : BOOL;
    Sequence : WORD;
    Sequence1 : WORD;
    Wait : TON;
END_VAR

IF Done THEN RETURN; END_IF;
Check := TRUE;
Ok := TRUE;
CASE Step OF
    0:
        全局变量_保持区.Store.dw签名 := 0;
        Runtime.w轴消费掩码 := 7;
        Runtime.b运行 := TRUE;
        Runtime.b待复位 := FALSE;
        Runtime.ast轴[0].b在线 := TRUE;
        Runtime.ast轴[0].b已使能 := TRUE;
        Runtime.ast轴[0].b静止 := TRUE;
        Runtime.ast轴[0].b可下发 := TRUE;
        Command[0] := XJV1_SIGNATURE_HI;
        Command[1] := XJV1_SIGNATURE_LO;
        Command[2] := 1;
        Server(Command := Command, Published := Published, Runtime := Runtime);
        Runtime.b待复位 := FALSE;
        Result := Axis_MoveToPoint(0, 120);
        Ok := NOT Result AND Axis状态(0).b错误 AND NOT Axis状态(0).b完成;
    1:
        Result := Axis_MoveToPoint(0, 16);
        Ok := Result AND Axis状态(0).b忙 AND NOT Axis状态(0).b完成;
        Result := Axis_Home(0);
        Ok := Ok AND NOT Result;
        (* 忙槽优先：无效新槽也不能改写已接受请求或其状态。 *)
        Result := Axis_MoveToPoint(0, 120);
        Ok := Ok AND NOT Result AND (全局变量_轴请求.ast请求[0].ui槽号 = 16)
            AND (全局变量_轴请求.ast请求[0].w命令 = 29)
            AND (全局变量_轴请求.ast请求[0].w错误 = 0);
    2:
        (* Free slot must reject through the real shared dispatch path. *)
        Command[2] := Command[2] + 1;
        Server(Command := Command, Published := Published, Runtime := Runtime);
        Ok := Axis状态(0).b错误 AND NOT Axis状态(0).b完成 AND (Runtime.aw轴命令[0] = 0);
    3:
        全局变量_保持区.Store.b已确认 := TRUE;
        全局变量_保持区.Store.aw点位[16, 0] := 0;
        全局变量_保持区.Store.aw点位[16, 1] := 1000;
        全局变量_保持区.Store.aw点位[16, 2] := 0;
        全局变量_保持区.Store.aw点位[16, 3] := 1000;
        全局变量_保持区.Store.aw点位[16, 4] := 3;
        Runtime.ast轴[0].w运动结果 := 2;
        Runtime.ast轴[0].w序列 := 65535;
        Result := Axis_MoveToPoint(0, 16);
        Ok := Result AND NOT Axis状态(0).b完成;
    4:
        Runtime.b待复位 := FALSE;
        Command[2] := Command[2] + 1;
        Server(Command := Command, Published := Published, Runtime := Runtime);
        Sequence := Runtime.aw轴序列[0];
        Manager(Runtime := Runtime);
        Ok := (Runtime.aw轴命令[0] = 27) AND (Sequence <> 65535)
            AND (Runtime.adi轴目标[0] = 1000) AND NOT Axis状态(0).b完成;
    5:
        Runtime.aw轴命令[0] := 0;
        Runtime.ast轴[0].w序列 := Sequence;
        Runtime.ast轴[0].w运动结果 := 1;
        Runtime.ast轴[0].b运动中 := TRUE;
        Runtime.ast轴[0].b静止 := FALSE;
        Manager(Runtime := Runtime);
        Ok := Axis状态(0).b忙 AND NOT Axis状态(0).b完成;
    6:
        Runtime.ast轴[0].w运动结果 := 2;
        Runtime.ast轴[0].b运动中 := FALSE;
        Runtime.ast轴[0].b静止 := TRUE;
        Manager(Runtime := Runtime);
        Ok := Axis状态(0).b完成 AND NOT Axis状态(0).b忙 AND NOT Axis状态(0).b错误;
    7:
        Result := Axis_MoveToPoint(0, 16);
        Ok := Result AND NOT Axis状态(0).b完成;
        Result := Axis_Stop(0);
        Ok := Ok AND Result AND NOT Axis状态(0).b完成 AND Axis状态(0).b错误
            AND (全局变量_轴请求.ast请求[0].w错误 = 19)
            AND (全局变量_轴请求.ast请求[0].w命令 = 26)
            AND NOT 全局变量_轴请求.ast请求[0].b已下发
            AND NOT 全局变量_轴请求.ast请求[0].b已接收;
    8:
        Command[2] := Command[2] + 1;
        Server(Command := Command, Published := Published, Runtime := Runtime);
        Manager(Runtime := Runtime);
        Ok := (Runtime.aw轴命令[0] = 26) AND NOT Axis状态(0).b完成;
    9:
        Result := Axis_Home(0);
        Runtime.b运行 := FALSE;
        Command[2] := Command[2] + 1;
        Server(Command := Command, Published := Published, Runtime := Runtime);
        Ok := Axis状态(0).b错误 AND (Runtime.aw轴命令[0] = 0);
    10:
        Ok := NOT Axis_MoveToPoint(16, 0) AND NOT Axis状态(16).b完成
            AND Axis状态(16).b错误 AND NOT Axis状态(16).b忙;
    11:
        Runtime.b运行 := TRUE;
        Runtime.ast轴[1].b在线 := TRUE;
        Runtime.ast轴[1].b已使能 := TRUE;
        Runtime.ast轴[1].b静止 := TRUE;
        Runtime.ast轴[1].b可下发 := TRUE;
        Result := Axis_Home(0);
        Ok := Result;
        Result := Axis_Home(1);
        Ok := Ok AND Result AND Axis状态(0).b忙 AND Axis状态(1).b忙;
    12:
        Command[2] := Command[2] + 1;
        Server(Command := Command, Published := Published, Runtime := Runtime);
        Sequence := Runtime.aw轴序列[0];
        Sequence1 := Runtime.aw轴序列[1];
        Ok := (Runtime.aw轴命令[0] = 22) AND (Runtime.aw轴命令[1] = 22);
    13:
        Runtime.ast轴[0].w序列 := Sequence;
        Runtime.ast轴[1].w序列 := Sequence1;
        Runtime.ast轴[0].w运动结果 := 1;
        Runtime.ast轴[1].w运动结果 := 1;
        Manager(Runtime := Runtime);
        Ok := Axis状态(0).b忙 AND Axis状态(1).b忙 AND NOT Axis状态(0).b完成 AND NOT Axis状态(1).b完成;
    14:
        Runtime.b暂停 := TRUE;
        Manager(Runtime := Runtime);
        Ok := Axis状态(0).b错误 AND Axis状态(1).b错误 AND NOT Axis状态(0).b完成 AND NOT Axis状态(1).b完成;
    15:
        Runtime.b暂停 := FALSE;
        Result := Axis_MoveToPoint(0, 16);
        Ok := Result;
        Command[3] := 26;
        Command[4] := 77;
        Command[5] := 16#0100;
        Command[2] := Command[2] + 1;
        Server(Command := Command, Published := Published, Runtime := Runtime);
        Ok := Ok AND (Runtime.aw轴命令[0] = 26) AND Axis状态(0).b错误 AND NOT Axis状态(0).b完成;
    16:
        Command[2] := Command[2] + 1;
        Server(Command := Command, Published := Published, Runtime := Runtime);
        Ok := (Runtime.aw轴命令[0] = 0) AND NOT Axis状态(0).b忙;
    17:
        Result := Axis_MoveToPoint(0, 16);
        Runtime.b暂停 := TRUE;
        Command[2] := Command[2] + 1;
        Server(Command := Command, Published := Published, Runtime := Runtime);
        Ok := Result AND Axis状态(0).b错误 AND (Runtime.aw轴命令[0] = 0);
    18:
        Runtime.b暂停 := FALSE;
        Runtime.b待复位 := TRUE;
        Result := Axis_Home(0);
        Command[2] := Command[2] + 1;
        Server(Command := Command, Published := Published, Runtime := Runtime);
        Ok := Result AND Axis状态(0).b错误 AND (Runtime.aw轴命令[0] = 0);
    19:
        (* Internal rejections must not replace the last network ACK. *)
        (* Wait past the 300ms publication period before checking network ACK. *)
        Wait(IN := TRUE, PT := T#400ms);
        Command[2] := Command[2] + 1;
        Server(Command := Command, Published := Published, Runtime := Runtime);
        IF NOT Wait.Q THEN Check := FALSE; RETURN; END_IF;
        Ok := (Published[3] = 77) AND (Published[4] = 0)
            AND (Published[5] = 16#0100) AND (Published[6] = 1);
        Done := TRUE;
END_CASE;
IF Check THEN
    IF Ok THEN Passed := Passed + 1;
    ELSE
        Failed := Failed + 1;
        IF FirstFailure = 0 THEN FirstFailure := Step + 1; END_IF;
    END_IF;
END_IF;
Step := Step + 1;
END_PROGRAM

(* ---- 程序_运行时自测.st ---- *)
(* Isolated simulator test. Fake feedback, no MC calls or physical outputs.
   Requires the xs_selftest isolated copy: lw已绑定气缸 is patched to 1,
   so cylinder 0 is bound and cylinder 1 stays unbound for these phases; the
   rated arrays are patched to 2147483647, which phase 25 depends on.
   Protocol 1.2: the official ModbusTCP slave writes the Holding image; this test
   writes the same Command array directly (payload first, SEQ last). *)
PROGRAM 程序_运行时自测
VAR
    st命令 : 类型_命令区;
    fb服务端 : 功能块_服务端;
    st发布 : 类型_发布区;
    st运行时 : 结构体_运行时;
    fb看门狗 : 功能块_看门狗;
    ui阶段 : UINT;
    i循环 : UINT;
    b正常 : BOOL;
    b检查 : BOOL;
    b提交 : BOOL;
    w命令码 : WORD;
    w对象字 : WORD;
    w序列 : WORD;
    w标记 : WORD;
    w结果 : WORD;
    udi通过 : UDINT;
    udi失败 : UDINT;
    ui首失败 : UINT;
    b完成 : BOOL;
END_VAR

IF b完成 THEN RETURN; END_IF;
b检查 := FALSE;
b提交 := FALSE;
b正常 := TRUE;
CASE ui阶段 OF
    0:
        全局变量_保持区.Store.dw签名 := 0;
        st运行时.b手动 := TRUE;
        st运行时.w轴消费掩码 := 7;
        FOR i循环 := 0 TO 2 DO
            st运行时.ast轴[i循环].b在线 := TRUE;
            st运行时.ast轴[i循环].b静止 := TRUE;
            st运行时.ast轴[i循环].b可下发 := TRUE;
        END_FOR;
        st命令[0] := XJV1_SIGNATURE_HI;
        st命令[1] := XJV1_SIGNATURE_LO;
    1:
        st命令[2] := 1;
    2:
        w命令码 := 20; w对象字 := 16#0100; b提交 := TRUE;
    3:
        b检查 := TRUE; b正常 := st运行时.aw轴命令[0] = 20;
    4:
        st运行时.ast轴[0].b已使能 := TRUE;
        st运行时.ast轴[0].b运动中 := TRUE;
        st运行时.ast轴[0].b静止 := FALSE;
        w命令码 := 21; b提交 := TRUE;
    5:
        b检查 := TRUE; b正常 := st运行时.aw轴命令[0] = 21;
    6:
        st运行时.ast轴[0].b运动中 := FALSE;
        st运行时.ast轴[0].b静止 := TRUE;
        w命令码 := 10; w对象字 := 0; b提交 := TRUE;
    7:
        b检查 := TRUE; b正常 := st运行时.b软急停 AND (st运行时.aw轴命令[0] = 26);
    8:
        w命令码 := 11; b提交 := TRUE;
    9:
        b检查 := TRUE; b正常 := NOT st运行时.b软急停 AND st运行时.b待复位;
    10:
        st运行时.ast轴[0].b故障 := TRUE;
        st运行时.ast轴[0].b静止 := FALSE;
        st运行时.ast轴[0].di速度 := 0;
        w命令码 := 1; b提交 := TRUE;
    11:
        b检查 := TRUE; b正常 := st运行时.b待复位 AND (st运行时.aw轴命令[0] = 26);
    12: ;
    13:
        b检查 := TRUE; b正常 := (st运行时.aw轴命令[0] = 23) AND (st运行时.aw轴序列[0] = w序列);
        FOR i循环 := 0 TO 2 DO
            st运行时.ast轴[i循环].b故障 := FALSE;
            st运行时.ast轴[i循环].b静止 := TRUE;
            st运行时.ast轴[i循环].w序列 := w序列;
            st运行时.ast轴[i循环].w运动结果 := 2;
        END_FOR;
    14:
        b检查 := TRUE; b正常 := NOT st运行时.b待复位;
    15:
        st运行时.aw轴命令[0] := 26;
        w结果 := 函数_动作许可(Code := 24, ObjectWord := 16#0100,
            HmiOnline := TRUE, JogBusy := FALSE, Resetting := FALSE,
            Runtime := st运行时, Store := 全局变量_保持区.Store);
        b检查 := TRUE; b正常 := w结果 = 10;
    16:
        w结果 := 函数_动作许可(Code := 26, ObjectWord := 16#0100,
            HmiOnline := FALSE, JogBusy := TRUE, Resetting := TRUE,
            Runtime := st运行时, Store := 全局变量_保持区.Store);
        b检查 := TRUE; b正常 := w结果 = 0;
    17:
        w结果 := 函数_动作许可(Code := 2, ObjectWord := 0,
            HmiOnline := TRUE, JogBusy := FALSE, Resetting := FALSE,
            Runtime := st运行时, Store := 全局变量_保持区.Store);
        b检查 := TRUE;
        IF 全局变量_运行配置.b正式流程已接入 THEN b正常 := w结果 = 0;
        ELSE b正常 := w结果 = 12;
        END_IF;
    18:
        st运行时.b硬急停 := TRUE;
        w结果 := 函数_动作许可(Code := 20, ObjectWord := 16#0100,
            HmiOnline := TRUE, JogBusy := FALSE, Resetting := FALSE,
            Runtime := st运行时, Store := 全局变量_保持区.Store);
        b检查 := TRUE; b正常 := w结果 = 3;
    19:
        st运行时.b硬急停 := FALSE;
        全局变量_保持区.Store.aw轴配置[0, 0] := 0;
        全局变量_保持区.Store.aw轴配置[0, 1] := 2000;
        全局变量_保持区.Store.aw轴配置[0, 2] := 0;
        全局变量_保持区.Store.aw轴配置[0, 3] := 1000;
        全局变量_保持区.Store.aw轴配置[0, 14] := 1;
        st运行时.ast轴[0].di位置 := 1500;
        w命令码 := 30; w对象字 := 16#0100; b提交 := TRUE;
    20:
        b检查 := TRUE; b正常 := st运行时.aw轴命令[0] = 0;
    21:
        st运行时.ast轴[0].b已使能 := FALSE;
        w结果 := 函数_动作许可(Code := 30, ObjectWord := 16#0100,
            HmiOnline := TRUE, JogBusy := FALSE, Resetting := FALSE,
            Runtime := st运行时, Store := 全局变量_保持区.Store);
        b检查 := TRUE; b正常 := w结果 = 6;
    22:
        (* 清故障在报警态必须可重试：残留的运动标志不再拒绝 23。 *)
        st运行时.ast轴[0].b运动中 := TRUE;
        w结果 := 函数_动作许可(Code := 23, ObjectWord := 16#0100,
            HmiOnline := TRUE, JogBusy := FALSE, Resetting := FALSE,
            Runtime := st运行时, Store := 全局变量_保持区.Store);
        b检查 := TRUE; b正常 := w结果 = 0;
    23:
        st运行时.ast轴[0].b运动中 := FALSE;
        st运行时.ast轴[0].b可下发 := FALSE;
        w结果 := 函数_动作许可(Code := 20, ObjectWord := 16#0100,
            HmiOnline := TRUE, JogBusy := FALSE, Resetting := FALSE,
            Runtime := st运行时, Store := 全局变量_保持区.Store);
        b检查 := TRUE; b正常 := w结果 = 10;
    24:
        st运行时.b硬急停 := TRUE;
        w结果 := 函数_动作许可(Code := 23, ObjectWord := 16#0100,
            HmiOnline := TRUE, JogBusy := FALSE, Resetting := FALSE,
            Runtime := st运行时, Store := 全局变量_保持区.Store);
        b检查 := TRUE; b正常 := w结果 = 3;
    25:
        st运行时.b硬急停 := FALSE;
        b检查 := TRUE;
        b正常 := NOT 函数_额定值(AxisIndex := 0, Field := 2, Value := 0)
            AND 函数_额定值(AxisIndex := 0, Field := 2, Value := 2147483647)
            AND NOT 函数_额定值(AxisIndex := 0, Field := 2, Value := 2147483648);
    26:
        b检查 := TRUE;
        b正常 := NOT 函数_额定值(AxisIndex := 16, Field := 2, Value := 1)
            AND NOT 函数_额定值(AxisIndex := 0, Field := 7, Value := 1);
    27:
        w命令码 := 42; w对象字 := 16#0201; b提交 := TRUE;
    28:
        b检查 := TRUE; b正常 := st运行时.aw气缸命令[1] = 0;
    29:
        w命令码 := 42; w对象字 := 16#0200; b提交 := TRUE;
    30:
        b检查 := TRUE; b正常 := (st运行时.aw气缸命令[0] = 42) AND (st运行时.aw气缸序列[0] = w序列);
    31:
        w命令码 := 40; w对象字 := 16#0200; b提交 := TRUE;
    32:
        b检查 := TRUE; b正常 := st运行时.aw气缸命令[0] = 0;
    33:
        w结果 := 函数_动作许可(Code := 42, ObjectWord := 16#0200,
            HmiOnline := FALSE, JogBusy := TRUE, Resetting := TRUE,
            Runtime := st运行时, Store := 全局变量_保持区.Store);
        b检查 := TRUE; b正常 := w结果 = 0;
    34:
        w结果 := 函数_动作许可(Code := 42, ObjectWord := 16#0201,
            HmiOnline := TRUE, JogBusy := FALSE, Resetting := FALSE,
            Runtime := st运行时, Store := 全局变量_保持区.Store);
        b检查 := TRUE; b正常 := w结果 = 4;
    35:
        fb看门狗(SignatureOK := TRUE, Heartbeat := 6);
    36:
        fb看门狗(SignatureOK := TRUE, Heartbeat := 7);
        b检查 := TRUE; b正常 := fb看门狗.Online;
    37:
        fb看门狗(SignatureOK := TRUE, Heartbeat := 7, StartJog := TRUE,
            StartObject := 16#0100, StartSequence := 9);
        b检查 := TRUE; b正常 := fb看门狗.JogActive;
    38:
        fb看门狗(SignatureOK := TRUE, Heartbeat := 7, StopJog := TRUE);
        b检查 := TRUE; b正常 := fb看门狗.CancelJog AND NOT fb看门狗.JogActive;
    39:
        (* Regression: a start pulse arriving while offline must establish and
           cancel the lease in the same scan instead of being dropped. *)
        fb看门狗(SignatureOK := FALSE, Heartbeat := 7, StartJog := TRUE,
            StartObject := 16#0100, StartSequence := 9);
        b检查 := TRUE; b正常 := fb看门狗.CancelJog AND NOT fb看门狗.JogActive;
    40:
        (* Drop the signature for one scan so the Server's own watchdogs go offline. *)
        w标记 := st运行时.aw轴序列[0];
        st命令[0] := 0;
    41:
        (* A command left in the Holding image across a reconnect is never
           replayed: on the connection edge the Server adopts its SEQ as the
           baseline. Code 26 is used because a stop bypasses every ordinary gate,
           so it would run here if the SEQ were treated as unconsumed. *)
        st命令[0] := XJV1_SIGNATURE_HI;
        w序列 := w序列 + 1;
        st命令[3] := 26;
        st命令[4] := w序列;
        st命令[5] := 16#0100;
    42:
        b检查 := TRUE; b正常 := st运行时.aw轴序列[0] = w标记;
    43:
        (* Positive control: the same payload under a genuinely new SEQ does run,
           so phase 42 can only pass because the SEQ was absorbed, not ignored. *)
        w命令码 := 26; w对象字 := 16#0100; b提交 := TRUE;
    44:
        b检查 := TRUE; b正常 := st运行时.aw轴序列[0] = w序列;
    45:
        st运行时.b硬急停 := FALSE;
        st运行时.b软急停 := TRUE;
        st运行时.b运行 := FALSE;
        st运行时.b待复位 := TRUE;
        w命令码 := 11; w对象字 := 0; b提交 := TRUE;
    46:
        b检查 := TRUE;
        b正常 := NOT st运行时.b软急停 AND NOT st运行时.b运行
            AND st运行时.b待复位;
    47:
        (* Clearing the software latch never restores motion permission:
           the axis is still not cleared for dispatch. *)
        w结果 := 函数_动作许可(Code := 20, ObjectWord := 16#0100,
            HmiOnline := TRUE, JogBusy := FALSE, Resetting := FALSE,
            Runtime := st运行时, Store := 全局变量_保持区.Store);
        b检查 := TRUE; b正常 := w结果 = 10;
    48:
        st运行时.b硬急停 := TRUE;
        st运行时.b软急停 := TRUE;
        w命令码 := 11; w对象字 := 0; b提交 := TRUE;
    49:
        b检查 := TRUE; b正常 := st运行时.b软急停 AND NOT st运行时.b运行;
    50:
        b完成 := TRUE;
END_CASE;
IF b检查 THEN
    IF b正常 THEN udi通过 := udi通过 + 1;
    ELSE
        udi失败 := udi失败 + 1;
        IF ui首失败 = 0 THEN ui首失败 := ui阶段; END_IF;
    END_IF;
END_IF;
IF b提交 THEN
    (* Same order as the host: payload words, then code, then SEQ last. *)
    FOR i循环 := 5 TO 31 DO st命令[i循环] := 0; END_FOR;
    st命令[5] := w对象字;
    st命令[3] := w命令码;
    w序列 := w序列 + 1;
    st命令[4] := w序列;
END_IF;
(* Heartbeat keeps the HMI online for the duration of the test. *)
st命令[2] := st命令[2] + 1;
fb服务端(Command := st命令, Published := st发布, Runtime := st运行时);
ui阶段 := ui阶段 + 1;
END_PROGRAM
